(* IEC 61131-3 sources: trust-platform/examples/OSCAT/compressor_pressure_filter/non-oop/src, 3 files *)

(* ---- Configuration.st ---- *)
CONFIGURATION CompressorPressureFilterClassicConfiguration
RESOURCE Cpu0 ON PLC
    TASK MainTask (INTERVAL := T#100ms, PRIORITY := 1);
    PROGRAM Main WITH MainTask : Main;
END_RESOURCE
END_CONFIGURATION

(* ---- Main.st ---- *)
PROGRAM Main
VAR
    PressureFilter : FT_PT1;
    PressureAlarm : HYST;
    RawPressureBar : REAL := REAL#11.0;
    FilteredPressureBar : REAL;
    AlarmActive : BOOL;
END_VAR

PressureFilter(in := RawPressureBar, T := T#1s, K := REAL#1.0);
FilteredPressureBar := PressureFilter.out;
PressureAlarm(In := FilteredPressureBar, HIGH_LIMIT := REAL#10.0, LOW_LIMIT := REAL#4.0);
AlarmActive := PressureAlarm.Q;
END_PROGRAM

(* ---- Tests.st ---- *)
TEST_PROGRAM CompressorPressureFilterClassicFiltersBeforeAlarm
VAR
    PressureFilter : FT_PT1;
    PressureAlarm : HYST;
END_VAR

PressureFilter(in := REAL#11.0, T := T#1s, K := REAL#1.0);
PressureAlarm(In := PressureFilter.out, HIGH_LIMIT := REAL#10.0, LOW_LIMIT := REAL#4.0);

ASSERT_NEAR(EXPECTED := REAL#11.0, ACTUAL := PressureFilter.out, DELTA := REAL#0.001);
ASSERT_TRUE(IN := PressureAlarm.Q);
END_TEST_PROGRAM
